INTERFACE I_Device

PROPERTY DeviceId : ST_DeviceId
GET
END_GET
END_PROPERTY

END_INTERFACE

(* stored: Version 1.1.0.1
   Itf I_Device: Id {33333333-3333-4333-8333-333333333333}
   Property DeviceId: Id {5e0ea2d3-5ebe-4720-9370-01c88b4afeb2}
   Get Get: Id {c595d6a1-ee48-4641-b1fb-ac450db55d1d} *)
